(* IEC 61131-3 sources: Antarbhukti-LLM/DatasetCreation/SeedSTs/batch2_filtered_NETWORK (part 4) *)

(* ---- TN_RECEIVE.ST ---- *)
(*@PROPERTIES_EX@
TYPE: POU
LOCALE: 0
IEC_LANGUAGE: ST
PLC_TYPE: independent
PROC_TYPE: independent
GROUP: TELNET_VISION
*)
(*@KEY@:DESCRIPTION*)
version 1.0		10. mai 2010
programmer		ks
tested by		ks

TN_RECEIVE empfängt Tastatureingaben vom Telnet Client und wertet diese aus

(*@KEY@:END_DESCRIPTION*)
FUNCTION_BLOCK TN_RECEIVE

(*Group:IN_OUT*)

VAR_IN_OUT
	R_BUF :	oscat_NETWORK_BUFFER;
	Xus_TN_SCREEN :	us_TN_SCREEN;
END_VAR

(*Group:lokal*)

VAR
	REQ_Size :	UINT;
	REQ1 :	BYTE;
	REQ2 :	BYTE;
	REQ3 :	BYTE;
END_VAR

(*@KEY@: WORKSHEET
NAME: TN_RECEIVE
IEC_LANGUAGE: ST
*)
(* -----------------------------------------------------------------*)
(* Datenempfang auswertung                                          *)
(* -----------------------------------------------------------------*)
Xus_TN_SCREEN.by_Input_ASCII_Code := BYTE#00;
Xus_TN_SCREEN.by_Input_Exten_Code := BYTE#00;

IF R_BUF.SIZE > UINT#0 THEN
  (* empfangene Daten auswerten *)
  REQ_Size := R_BUF.SIZE;
  REQ1 := R_BUF.BUFFER[0];
  REQ2 := R_BUF.BUFFER[1];
  REQ3 := R_BUF.BUFFER[2];

  IF REQ1 = BYTE#27 AND REQ_Size >= UINT#3 THEN (* Escape *)
    IF REQ2 = BYTE#91 THEN (* Cursor code *)
      IF (REQ3 >= BYTE#65 AND REQ3 <= BYTE#68) OR (REQ3 = BYTE#72) OR (REQ3 = BYTE#75) THEN (* 65..68 = Cursor o,u,r,l / 72 = POS1 / 75 = ENDE *)
        Xus_TN_SCREEN.by_Input_Exten_Code := REQ3;
      END_IF;
    ELSIF REQ2 = BYTE#79 THEN (* Sondertasten F1/F2/F3/F4 *)
      IF REQ3 >= BYTE#80 AND REQ3 <= BYTE#83 THEN
        Xus_TN_SCREEN.by_Input_Exten_Code := REQ3;
      END_IF;
    END_IF;
  ELSIF REQ1 >= BYTE#32 AND REQ1 <= BYTE#126 THEN
	Xus_TN_SCREEN.by_Input_ASCII_Code := REQ1;
    Xus_TN_SCREEN.bo_Input_ASCII_IsNum := ISC_NUM(REQ1); (* Auswertung auf Zahleneingabe *)
  ELSIF REQ1 = BYTE#8 OR REQ1 = BYTE#9 OR REQ1 = BYTE#13 OR REQ1 = BYTE#27 THEN (* prüfe auf Steuerzeichen 8=Backspace / 9=Tabulator / 13=Return / 27=Escape *)
	Xus_TN_SCREEN.by_Input_Exten_Code := REQ1;
  END_IF;

  (* Empfangsbuffer Datenlänge null eintragen (Telegramm zerstören *)
  R_BUF.SIZE := UINT#00;
END_IF;

(* revision history
ks	10. mai. 2010	rev 1.0
	original version
*)

(*@KEY@: END_WORKSHEET *)
END_FUNCTION_BLOCK

(* ---- WORLD_WEATHER.ST ---- *)
(*@PROPERTIES_EX@
TYPE: POU
LOCALE: 0
IEC_LANGUAGE: ST
PLC_TYPE: independent
PROC_TYPE: independent
GROUP: WEATHER
*)
(*@KEY@:DESCRIPTION*)
version 1.3		05. jan 2012
programmer 		ks
tested by		ks

WORLD_WEATHER lädt von worldweather.com eine Wetter csv-datei und analysiert die Daten und legt diese in einem Array ab
Die Wetterdaten werden für 5 tage aufbereitet

(*@KEY@:END_DESCRIPTION*)
FUNCTION_BLOCK WORLD_WEATHER

(*Group:in_out*)

VAR_INPUT
	ACTIVATE :	BOOL;
	LATITUDE :	REAL;
	LONGITUDE :	REAL;
	KEY :	oscat_STRING30;
END_VAR

VAR_OUTPUT
	BUSY :	BOOL;
	DONE :	BOOL;
	ERROR_C :	DWORD;
	ERROR_T :	BYTE;
END_VAR

VAR_IN_OUT
	IP_C :	oscat_IP_C;(*IP_Control Verwaltungsstruktur*)
	S_BUF :	oscat_NETWORK_BUFFER;
	R_BUF :	oscat_NETWORK_BUFFER;
	WW :	oscat_WORLD_WEATHER_DATA;
END_VAR

(*Group:var*)

VAR
	CHK_REAL :	CHK_REAL;
	REAL_TO_STRF :	REAL_TO_STRF;
	URL_DATA :	oscat_url;
	DNS_CLIENT :	DNS_CLIENT;
	HTTP_GET :	HTTP_GET;
	CPB :	CSV_PARSER_BUF;
	STRING_TO_URL :	STRING_TO_URL;
	FLOAT_TO_REAL :	FLOAT_TO_REAL;
	last_state :	BOOL;
	value_int :	INT;
	value_real :	REAL;
	v_real :	REAL;
	state :	INT;
	url_str :	oscat_STRING250;
	offset :	UDINT;
	size :	INT;
	sep :	BYTE;
	cnt :	INT;
	day :	INT;
	idx :	INT;
	run :	BYTE;
	result :	BYTE;
	value :	oscat_STRING250;
	DEC_TO_INT :	DEC_TO_INT;
	pos :	INT;
END_VAR

(*@KEY@: WORKSHEET
NAME: WORLD_WEATHER
IEC_LANGUAGE: ST
*)
CASE state OF

00:
	IF ACTIVATE AND NOT last_state THEN
		state := 20;
		DONE := FALSE;
		BUSY := TRUE;
		ERROR_C := DWORD#0;
		ERROR_T := BYTE#0;
	END_IF;

20: (* URL for DNS UND HTTP-GET *)
	(* Example: http://free.worldweatheronline.com/feed/weather.ashx?q=48.21,16.37&format=csv&num_of_days=5&key=xxxxxxxxxxxxxxxxxxxxxx *)

	REAL_TO_STRF(IN:=LATITUDE,N:=6,D:='.');
	url_str := CONCAT('http://free.worldweatheronline.com/feed/weather.ashx?q=',REAL_TO_STRF.REAL_TO_STRF);
	url_str := CONCAT(url_str,',');
	REAL_TO_STRF(IN:=LONGITUDE,N:=6,D:='.');
	url_str := CONCAT(url_str,REAL_TO_STRF.REAL_TO_STRF);
	url_str := CONCAT(url_str,'&format=csv&num_of_days=5&key=');
	url_str := CONCAT(url_str,key);

	STRING_TO_URL(STR:=url_str, DEFAULT_PROTOCOL:='', DEFAULT_PATH:='' );
  	URL_DATA:=STRING_TO_URL.STRING_TO_URL;

	state := 40;

40:
	IF DNS_CLIENT.DONE THEN
		state := 60;
	ELSIF (DNS_CLIENT.ERROR > DWORD#00) THEN
		(* Fehlerbehandlung *)
		ERROR_C := DNS_CLIENT.ERROR;
		ERROR_T := BYTE#01;
		state   := 100;
	END_IF;

60:
	IF HTTP_GET.DONE THEN
		sep := BYTE#0;
		idx := 0;
		day := 0;
		cnt := 0;
		OFFSET := UINT_TO_UDINT(HTTP_GET.BODY_START); (* Start Offset vorgeben *)
		size := UINT_TO_INT(HTTP_GET.BODY_STOP); (* End Position *)
		run := BYTE#1; (* Element suchen *)
		state := 80;

	ELSIF (HTTP_GET.ERROR > DWORD#00) THEN
		(* Fehlerbehandlung *)
		ERROR_C := HTTP_GET.ERROR;
		ERROR_T := BYTE#02;
		state := 100;
	END_IF;

80:	IF run = BYTE#0 THEN (* kein Befehl mehr aktiv ? *)
		run := BYTE#1; (*  nächstes Element suchen  *)
		IF result = BYTE#1 OR result = BYTE#2 THEN
			value_int := 0;
			value_real := 0.0;
			(* automatische konvertierung in real und int ausführen *)
			IF LEN(value) <= 20 THEN
      			FLOAT_TO_REAL(FLT:=value);
				v_real := FLOAT_TO_REAL.FLOAT_TO_REAL;
				CHK_REAL(X := v_real); (* !!! prüft auf gültigen REAL Wert, ansonsten stürzt Twincat ab !!!!  *)
				IF CHK_REAL.CHK_REAL = BYTE#0 THEN
					value_real := v_real;
					value_int := REAL_TO_INT(value_real);
				END_IF;
			END_IF;
			cnt := cnt + 1;
			IF cnt >=8 AND cnt <= 87 THEN
				IF cnt > 22 THEN
					CASE idx OF
					00:	WW.DAY[day].DATE_OF_DAY := value;
					01:	WW.DAY[day].TEMP_MAX_C := value_int;
					02:	WW.DAY[day].TEMP_MAX_F := value_int;
					03:	WW.DAY[day].TEMP_MIN_C := value_int;
					04:	WW.DAY[day].TEMP_MIN_F := value_int;
					05:	WW.DAY[day].WIND_SPEED_MILES := value_int;
					06:	WW.DAY[day].WIND_SPEED_KMPH := value_int;
					07:	WW.DAY[day].WIND_DIR_DEGREE := value_int;
					08:	WW.DAY[day].WIND_DIR16POINT := value;
					09:	WW.DAY[day].WEATHER_CODE := value_int;
					10:	pos := FIND(value, '/wsymbol_');
                        IF pos > 0 AND LEN(value) > pos + 13 THEN
                            DEC_TO_INT(DEC:=MID(value,4,pos + 9));
                            WW.DAY[day].WEATHER_ICON := DEC_TO_INT.DEC_TO_INT;
                        ELSE
       						WW.DAY[day].WEATHER_ICON := 0;
                        END_IF;
					11:	WW.DAY[day].WEATHER_DESC := value;
					12:	WW.DAY[day].PRECIPMM := value_real;
					END_CASE;
					idx := idx + 1;
					IF idx > 12 THEN
						idx := 0;
						day := day + 1;
					END_IF;
				ELSE
					CASE cnt OF
					08:	sep := BYTE#44; (* ab jetzt mit Trennzeichen arbeiten, *)
					09:	WW.CUR.OBSERVATION_TIME := value;
					10:	WW.CUR.TEMP_C := value_int;
					11:	WW.CUR.WEATHER_CODE := value_int;
					12:	pos := FIND(value, '/wsymbol_');
                        IF pos > 0 AND LEN(value) > pos + 13 THEN
                            DEC_TO_INT(DEC:=MID(value,4,pos + 9));
                            WW.CUR.WEATHER_ICON := DEC_TO_INT.DEC_TO_INT;
                        ELSE
       						WW.CUR.WEATHER_ICON := 0;
                        END_IF;
					13:	WW.CUR.WEATHER_DESC := value;
					14:	WW.CUR.WIND_SPEED_MILES := value_int;
					15:	WW.CUR.WIND_SPEED_KMPH := value_int;
					16:	WW.CUR.WIND_DIR_DEGREE := value_int;
					17:	WW.CUR.WIND_DIR16POINT := value;
					18:	WW.CUR.PRECIPMM := value_real;
					19:	WW.CUR.HUMIDITY := value_int;
					20:	WW.CUR.VISIBILITY := value_int;
					21:	WW.CUR.PRESSURE := value_int;
					22:	WW.CUR.CLOUDOVER := value_int;
					END_CASE;
				END_IF;
			END_IF;
		ELSIF result = BYTE#10 THEN (* nichts mehr gefunden *)
			DONE  := TRUE;
			run := BYTE#0; (* Auswertung beenden *)
			state := 100;
		END_IF;
	END_IF;

100:
	(* UNLOCK HTTP DATA *)
	IF (NOT HTTP_GET.DONE) THEN
		state := 0;
		BUSY := FALSE;
		DONE := ERROR_T = BYTE#0;
	END_IF;

END_CASE;

(* ---------------- DNS --------------- *)
DNS_CLIENT.IP_C     := IP_C;
DNS_CLIENT.S_BUF    := S_BUF;
DNS_CLIENT.R_BUF    := R_BUF;
DNS_CLIENT.DOMAIN   := URL_DATA.DOMAIN;
DNS_CLIENT.IP4_DNS  := DWORD#00;
DNS_CLIENT.ACTIVATE := state=40; (* DNS Start *)
DNS_CLIENT();
IP_C  := DNS_CLIENT.IP_C;
S_BUF := DNS_CLIENT.S_BUF;
R_BUF := DNS_CLIENT.R_BUF;

(* nicht oder nicht direkt verwendete Parameter *)
(* DWORD :=DNS_CLIENT.IP4;
   BOOL  :=DNS_CLIENT.DONE;
   BYTE  :=DNS_CLIENT.ERROR; *)
(* -------------------------------------*)

(* ------------- HTTP_GET --------------- *)

HTTP_GET.IP_C        := IP_C;
HTTP_GET.S_BUF       := S_BUF;
HTTP_GET.R_BUF       := R_BUF;
HTTP_GET.IP4         := DNS_CLIENT.IP4;
HTTP_GET.GET         := state=60;
HTTP_GET.MODE        := BYTE#2; (* HTTP 1.1 mit persistenter Verbindung *)
HTTP_GET.UNLOCK_BUF  := state=100;
HTTP_GET.URL_DATA    := URL_DATA;
HTTP_GET();
IP_C     := HTTP_GET.IP_C;
S_BUF    := HTTP_GET.S_BUF;
R_BUF    := HTTP_GET.R_BUF;
URL_DATA := HTTP_GET.URL_DATA;

(* nicht oder nicht direkt verwendete Parameter *)
(*STRING := HTTP_GET.HTTP_STATUS;
  UINT :=HTTP_GET.HEADER_START;
  UINT :=HTTP_GET.HEADER_STOP;
  UINT :=HTTP_GET.BODY_START;
  UINT :=HTTP_GET.BODY_STOP;
  BOOL :=HTTP_GET.DONE;
  BYTE :=HTTP_GET.ERROR;
*)
(* -------------------------------------*)

CPB(SEP:=sep,RUN:=run,OFFSET:=offset,VALUE:=value,PT:=R_BUF); (* CSV PARAMETER BUF *)
run:=CPB.RUN;
offset:=CPB.OFFSET;
value:=CPB.VALUE;
R_BUF:=CPB.PT;
result:=CPB.RESULT;

last_state := ACTIVATE;

(* revision history
ks	01.oct. 2010	rev 1.0
	original version

ks	01.feb. 2011	rev 1.1
	rücksetzen von cnt

ks	07.apr. 2011	rev 1.2
	neue Domain "free.worldweatheronline.com" (Ab 30.04.2011 notwendig)

ks	05.jan. 2012	rev 1.3
	neues datenelement "icon" integriert, REAL_TO_STRF parameter D
*)

(*@KEY@: END_WORKSHEET *)
END_FUNCTION_BLOCK

(* ---- YAHOO_WEATHER.ST ---- *)
(*@PROPERTIES_EX@
TYPE: POU
LOCALE: 0
IEC_LANGUAGE: ST
PLC_TYPE: independent
PROC_TYPE: independent
GROUP: WEATHER
*)
(*@KEY@:DESCRIPTION*)

version 1.3		04. may. 2011
programmer 		ks
tested by		ks

YAHOO_WEATHER lädt vom Yahoo-Webserver einen Wetter RSS-Feed und analysiert die Daten und legt diese in einem Array ab
(*@KEY@:END_DESCRIPTION*)
FUNCTION_BLOCK YAHOO_WEATHER

(*Group:in_out*)

VAR_IN_OUT
	IP_C :	oscat_IP_C;(*IP_Control Verwaltungsstruktur*)
	S_BUF :	oscat_NETWORK_BUFFER;
	R_BUF :	oscat_NETWORK_BUFFER;
	YW :	oscat_YAHOO_WEATHER_DATA;
END_VAR

VAR_INPUT
	ACTIVATE :	BOOL;
	UNITS :	BOOL;
	LOCATION :	oscat_STRING20;
END_VAR

VAR_OUTPUT
	BUSY :	BOOL;
	DONE :	BOOL;
	ERROR_C :	DWORD;
	ERROR_T :	BYTE;
END_VAR

(*Group:var*)

VAR
	CTRL :	oscat_XML_CONTROL;
	XML_READER :	XML_READER;
	URL_DATA :	oscat_url;
	DNS_CLIENT :	DNS_CLIENT;
	STRING_TO_URL :	STRING_TO_URL;
	HTTP_GET :	HTTP_GET;
	FLOAT_TO_REAL :	FLOAT_TO_REAL;
	CHK_REAL :	CHK_REAL;
	last_state :	BOOL;
	value_int :	INT;
	value_real :	REAL;
	v_real :	REAL;
	state :	INT;
END_VAR

(*@KEY@: WORKSHEET
NAME: YAHOO_WEATHER
IEC_LANGUAGE: ST
*)

CASE state OF

00:
  IF ACTIVATE AND NOT last_state THEN
    state := 20;
	DONE := FALSE;
	BUSY := TRUE;
	ERROR_C := DWORD#0;
	ERROR_T := BYTE#0;
  END_IF;

20: (* URL for DNS UND HTTP-GET *)
  (* Example: http://weather.yahooapis.com/forecastrss?p=94089&u=c *)
  STRING_TO_URL.STR:='http://weather.yahooapis.com/forecastrss';
  STRING_TO_URL.DEFAULT_PROTOCOL:='';
  STRING_TO_URL.DEFAULT_PATH:='';
  STRING_TO_URL();
  URL_DATA:=STRING_TO_URL.STRING_TO_URL;

  URL_DATA.QUERY := CONCAT('w=',LOCATION);

  IF UNITS THEN
    URL_DATA.QUERY := CONCAT(URL_DATA.QUERY,'&u=f'); (* fahrenheit *)
  ELSE
    URL_DATA.QUERY := CONCAT(URL_DATA.QUERY,'&u=c'); (* celsius *)
  END_IF;

  state := 40;

40:
  IF DNS_CLIENT.DONE THEN
    state := 60;
  ELSIF (DNS_CLIENT.ERROR > DWORD#00) THEN
    (* Fehlerbehandlung *)
    ERROR_C := DNS_CLIENT.ERROR;
	ERROR_T := BYTE#01;
    state   := 100;
  END_IF;

60:
  IF HTTP_GET.DONE THEN
    state := 80;
    CTRL.START_POS := HTTP_GET.BODY_START;
    CTRL.STOP_POS  := HTTP_GET.BODY_STOP;
    CTRL.COMMAND   := WORD#2#10000000_00011000; (* ONLY TEXT AND ATTRIBUTE *)
	CTRL.WATCHDOG  := T#1ms;

  ELSIF (HTTP_GET.ERROR > DWORD#00) THEN
    (* Fehlerbehandlung *)
    ERROR_C := HTTP_GET.ERROR;
	  ERROR_T := BYTE#02;
    state   := 100;
  END_IF;

80:
  (* XML Daten seriell lesen *)
  XML_READER.CTRL := CTRL;
  XML_READER.BUF  := R_BUF.BUFFER;
  XML_READER();
  CTRL         := XML_READER.CTRL;
  R_BUF.BUFFER := XML_READER.BUF;

  IF CTRL.TYP < 98 THEN (* nur auswerten wenn kein Watchdog durchlauf *)
    value_int := 0;
	value_real := 0.0;
	(* automatische konvertierung in real und int ausführen *)
	IF LEN(CTRL.VALUE) <= 20 THEN
      FLOAT_TO_REAL(FLT:=CTRL.VALUE);
      v_real:=FLOAT_TO_REAL.FLOAT_TO_REAL;
	  CHK_REAL(X:= v_real); (* !!! prüft auf gültigen REAL Wert, ansonsten stürzt Twincat ab !!!!  *)
	  IF CHK_REAL.CHK_REAL = BYTE#0 THEN
	    value_real := v_real;
		value_int := REAL_TO_INT(value_real);
	  END_IF;
	END_IF;

    IF CTRL.COUNT < UINT#52 THEN (* Performance-Teilung *)
      (* ------------ Teil 1 --------------*)
      CASE UINT_TO_INT(CTRL.COUNT) OF
        027: YW.TimeToLive := value_int;
        030: YW.location_city := CTRL.VALUE;
        031: YW.location_region := CTRL.VALUE;
        032: YW.location_country := CTRL.VALUE;
        035: YW.unit_temperature := CTRL.VALUE;
        036: YW.unit_distance := CTRL.VALUE;
        037: YW.unit_pressure := CTRL.VALUE;
        038: YW.unit_speed := CTRL.VALUE;
        041: YW.wind_chill := value_int;
        042: YW.wind_direction := value_int;
        043: YW.wind_speed := value_real;
        046: YW.atmosphere_humidity := value_int;
        047: YW.atmosphere_visibility := value_real;
        048: YW.atmosphere_pressure := value_int;
        049: YW.atmosphere_rising := value_int;
      END_CASE;
    ELSE
      (* ------------ Teil 2 --------------*)
      CASE UINT_TO_INT(CTRL.COUNT) OF
        052: YW.astronomy_sunrise := CTRL.VALUE;
        053: YW.astronomy_sunset := CTRL.VALUE;
        077: YW.geo_latitude := value_real;
        080: YW.geo_longitude := value_real;
        089: YW.cur_conditions_text := CTRL.VALUE;
		090: YW.cur_conditions_code := value_int;
			 YW.cur_conditions_icon := value_int;
        091: YW.cur_conditions_temp := value_int;
        100: YW.forcast_today_low_temp := value_int;
        101: YW.forcast_today_high_temp := value_int;
        102: YW.forcast_today_text := CTRL.VALUE;
		103: YW.forcast_today_code := value_int;
			 YW.forcast_today_icon := value_int;
        108: YW.forcast_tomorrow_low_temp := value_int;
        109: YW.forcast_tomorrow_high_temp := value_int;
        110: YW.forcast_tomorrow_text := CTRL.VALUE;
		111: YW.forcast_tomorrow_code := value_int;
			 YW.forcast_tomorrow_icon := value_int;
      END_CASE;
    END_IF;
  ELSIF CTRL.TYP = 99 THEN (* EXIT - letztes Element gelesen *)
    DONE  := TRUE;
    state := 100;
  END_IF;

100:
  (* UNLOCK HTTP DATA *)
  IF (NOT HTTP_GET.DONE) THEN
    state := 0;
    BUSY  := FALSE;
    DONE := ERROR_T = BYTE#0;
  END_IF;

END_CASE;

(* ---------------- DNS --------------- *)
DNS_CLIENT.IP_C     := IP_C;
DNS_CLIENT.S_BUF    := S_BUF;
DNS_CLIENT.R_BUF    := R_BUF;
DNS_CLIENT.DOMAIN   := URL_DATA.DOMAIN;
DNS_CLIENT.IP4_DNS  := DWORD#00;
DNS_CLIENT.ACTIVATE := state=40; (* DNS Start *)
DNS_CLIENT();
IP_C  := DNS_CLIENT.IP_C;
S_BUF := DNS_CLIENT.S_BUF;
R_BUF := DNS_CLIENT.R_BUF;

(* nicht oder nicht direkt verwendete Parameter *)
(* DWORD :=DNS_CLIENT.IP4;
   BOOL  :=DNS_CLIENT.DONE;
   BYTE  :=DNS_CLIENT.ERROR; *)
(* -------------------------------------*)

(* ------------- HTTP_GET --------------- *)

HTTP_GET.IP_C        := IP_C;
HTTP_GET.S_BUF       := S_BUF;
HTTP_GET.R_BUF       := R_BUF;
HTTP_GET.IP4         := DNS_CLIENT.IP4;
HTTP_GET.GET         := state=60;
HTTP_GET.MODE        := BYTE#2; (* HTTP 1.1 mit persistenter Verbindung *)
HTTP_GET.UNLOCK_BUF  := state=100;
HTTP_GET.URL_DATA    := URL_DATA;
HTTP_GET();
IP_C     := HTTP_GET.IP_C;
S_BUF    := HTTP_GET.S_BUF;
R_BUF    := HTTP_GET.R_BUF;
URL_DATA := HTTP_GET.URL_DATA;

(* nicht oder nicht direkt verwendete Parameter *)
(*STRING := HTTP_GET.HTTP_STATUS;
  UINT :=HTTP_GET.HEADER_START;
  UINT :=HTTP_GET.HEADER_STOP;
  UINT :=HTTP_GET.BODY_START;
  UINT :=HTTP_GET.BODY_STOP;
  BOOL :=HTTP_GET.DONE;
  BYTE :=HTTP_GET.ERROR;
*)
(* -------------------------------------*)

last_state := ACTIVATE;

(* revision history
ks	18. dez. 2008	rev 1.0
	original version

ks	01. oct. 2009	rev 1.1
	YAHOO_WEATHER_DATA

ks	24. sep. 2010	rev 1.2
	new URL-Location-parameter and REAL_CHECK (TwinCat BUG)

ks	04. may. 2011	rev 1.3
	neue elemente:  CUR_CONDITIONS_ICON, FORCAST_TODAY_ICON, FORCAST_TOMORROW_ICON

*)

(*@KEY@: END_WORKSHEET *)
END_FUNCTION_BLOCK
